// TIA Portal V20 export
// export: Created 2026-10-19T18:02:13.1059289Z, ExportSetting WithDefaults, DisplayName Totally Integrated Automation Portal, DisplayVersion V20 Update 6, DisplayName TIA Portal Openness, DisplayVersion V20 Update 6, DisplayName TIA Portal Version Control Interface, DisplayVersion V20 Update 6, DisplayName SINAMICS Startdrive Advanced, DisplayVersion V20 SP1, DisplayName SINAMICS Startdrive G130, G150, S120, S150, SINAMICS MV, G220, S200, S210, DisplayVersion V20 SP1, DisplayName SINAMICS Startdrive G110M, G120, G120C, G120D, G120P, G115D, DisplayVersion V20 SP1, DisplayName STEP 7 Professional, DisplayVersion V20 Update 6, DisplayName STEP 7 Safety, DisplayVersion V20 Update 2, DisplayName WinCC Basic/Comfort/Advanced, DisplayVersion V20 Update 6, DisplayName WinCC Unified, DisplayVersion V20 Update 6
FUNCTION "REMOTE PANEL" : Void   // FC1, F_LAD
{ S7_Optimized_Access := 'TRUE' }
VERSION : 0.1
// stored: AutoNumber true, IsIECCheckEnabled false, UDAEnableTagReadback false
   VAR_INPUT
      ACK : Bool;
   END_VAR
   VAR_OUTPUT
      OK : Bool;
      ESTOP_INBOUND : Bool;
   END_VAR
BEGIN

REGION Network 1: REMOTE PANEL OK
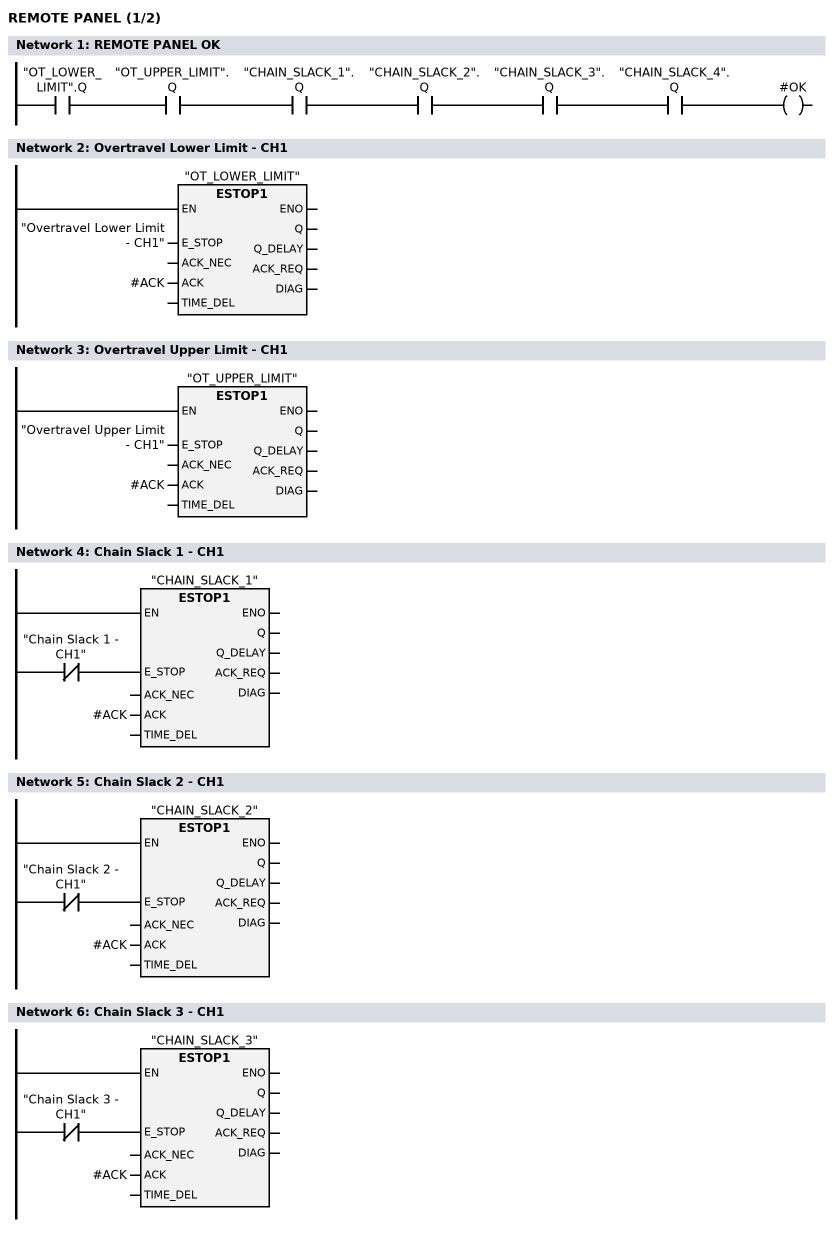
   RUNG wire#powerrail
      Contact( "OT_LOWER_LIMIT".Q )
      Contact( "OT_UPPER_LIMIT".Q )
      Contact( "CHAIN_SLACK_1".Q )
      Contact( "CHAIN_SLACK_2".Q )
      Contact( "CHAIN_SLACK_3".Q )
      Contact( "CHAIN_SLACK_4".Q )
      Coil( #OK )
   END_RUNG
   // the same network as SCL:
   #OK := "OT_LOWER_LIMIT".Q AND "OT_UPPER_LIMIT".Q AND "CHAIN_SLACK_1".Q AND "CHAIN_SLACK_2".Q AND "CHAIN_SLACK_3".Q AND "CHAIN_SLACK_4".Q;
END_REGION

REGION Network 2: Overtravel Lower Limit - CH1
   RUNG wire#powerrail
      "OT_LOWER_LIMIT".ESTOP1(E_STOP := "Overtravel Lower Limit - CH1", ACK_NEC :=, ACK := #ACK, TIME_DEL :=, Q =>, Q_DELAY =>, ACK_REQ =>, DIAG =>)
   END_RUNG
   // the same network as SCL:
   "OT_LOWER_LIMIT"(E_STOP := "Overtravel Lower Limit - CH1", ACK := #ACK);   // ESTOP1
END_REGION

REGION Network 3: Overtravel Upper Limit - CH1
   RUNG wire#powerrail
      "OT_UPPER_LIMIT".ESTOP1(E_STOP := "Overtravel Upper Limit - CH1", ACK_NEC :=, ACK := #ACK, TIME_DEL :=, Q =>, Q_DELAY =>, ACK_REQ =>, DIAG =>)
   END_RUNG
   // the same network as SCL:
   "OT_UPPER_LIMIT"(E_STOP := "Overtravel Upper Limit - CH1", ACK := #ACK);   // ESTOP1
END_REGION

REGION Network 4: Chain Slack 1 - CH1
   RUNG wire#powerrail
      "CHAIN_SLACK_1".ESTOP1(E_STOP := wire#w1, ACK_NEC :=, ACK := #ACK, TIME_DEL :=, Q =>, Q_DELAY =>, ACK_REQ =>, DIAG =>)
   END_RUNG
   RUNG wire#powerrail
      I_Contact( "Chain Slack 1 - CH1" )
   END_RUNG wire#w1
   // the same network as SCL:
   "CHAIN_SLACK_1"(E_STOP := NOT "Chain Slack 1 - CH1", ACK := #ACK);   // ESTOP1
END_REGION

REGION Network 5: Chain Slack 2 - CH1
   RUNG wire#powerrail
      "CHAIN_SLACK_2".ESTOP1(E_STOP := wire#w1, ACK_NEC :=, ACK := #ACK, TIME_DEL :=, Q =>, Q_DELAY =>, ACK_REQ =>, DIAG =>)
   END_RUNG
   RUNG wire#powerrail
      I_Contact( "Chain Slack 2 - CH1" )
   END_RUNG wire#w1
   // the same network as SCL:
   "CHAIN_SLACK_2"(E_STOP := NOT "Chain Slack 2 - CH1", ACK := #ACK);   // ESTOP1
END_REGION

REGION Network 6: Chain Slack 3 - CH1
   RUNG wire#powerrail
      "CHAIN_SLACK_3".ESTOP1(E_STOP := wire#w1, ACK_NEC :=, ACK := #ACK, TIME_DEL :=, Q =>, Q_DELAY =>, ACK_REQ =>, DIAG =>)
   END_RUNG
   RUNG wire#powerrail
      I_Contact( "Chain Slack 3 - CH1" )
   END_RUNG wire#w1
   // the same network as SCL:
   "CHAIN_SLACK_3"(E_STOP := NOT "Chain Slack 3 - CH1", ACK := #ACK);   // ESTOP1
END_REGION

REGION Network 7: Chain Slack 4 - CH1
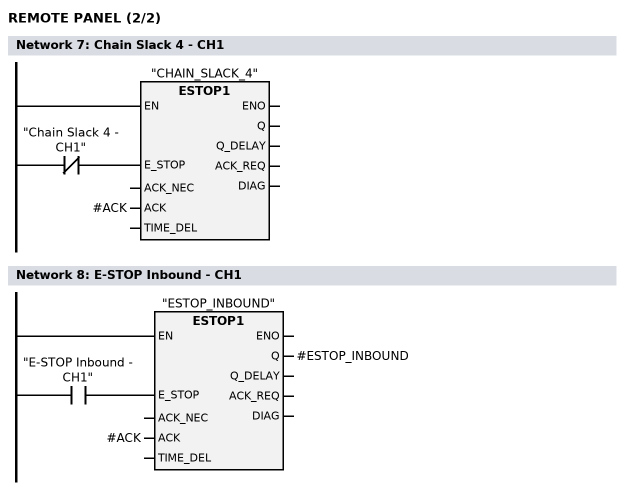
   RUNG wire#powerrail
      "CHAIN_SLACK_4".ESTOP1(E_STOP := wire#w1, ACK_NEC :=, ACK := #ACK, TIME_DEL :=, Q =>, Q_DELAY =>, ACK_REQ =>, DIAG =>)
   END_RUNG
   RUNG wire#powerrail
      I_Contact( "Chain Slack 4 - CH1" )
   END_RUNG wire#w1
   // the same network as SCL:
   "CHAIN_SLACK_4"(E_STOP := NOT "Chain Slack 4 - CH1", ACK := #ACK);   // ESTOP1
END_REGION

REGION Network 8: E-STOP Inbound - CH1
   RUNG wire#powerrail
      "ESTOP_INBOUND".ESTOP1(E_STOP := wire#w1, ACK_NEC :=, ACK := #ACK, TIME_DEL :=, Q => #ESTOP_INBOUND, Q_DELAY =>, ACK_REQ =>, DIAG =>)
   END_RUNG
   RUNG wire#powerrail
      Contact( "E-STOP Inbound - CH1" )
   END_RUNG wire#w1
   // the same network as SCL:
   "ESTOP_INBOUND"(E_STOP := "E-STOP Inbound - CH1", ACK := #ACK, Q => #ESTOP_INBOUND);   // ESTOP1
END_REGION
END_FUNCTION
